{attribute 'Tc2GvlVarNames'}
VAR_GLOBAL
	(*fbCheckArrayBounds: FB_CheckArrayBounds;*)

END_VAR

(* stored: Version 1.1.0.1, ProductVersion 3.1.4024.15
   GVL GVL_FB_CheckArrayBounds: Id {ec733504-a7f4-4530-b80e-c4be2bffa9a9} *)
